(* IEC 61131-3 sources: codesys/project-view/Device/Plc Logic/Application/00-封装FC/DATA类型转换, 14 files *)

(* ---- FC_1DINT_TO_1DWORD.st ---- *)
FUNCTION FC_1DINT_TO_1DWORD : DWORD
VAR_INPUT
	diIN:DINT;
END_VAR
VAR
	pdw:POINTER TO DWORD;
END_VAR
// --- implementation ---
pdw:=ADR(diIN);
FC_1DINT_TO_1DWORD:=pdw^;
END_FUNCTION

(* ---- FC_1DWORD_TO_1REAL.st ---- *)
FUNCTION FC_1DWORD_TO_1REAL : REAL
VAR_INPUT
	dwIN:DWORD;
END_VAR
VAR
	pr:POINTER TO REAL;
END_VAR
// --- implementation ---
pr:=ADR(dwIN);
FC_1DWORD_TO_1REAL:=pr^;
END_FUNCTION

(* ---- FC_1REAL_TO_1DWORD.st ---- *)
FUNCTION FC_1REAL_TO_1DWORD : DWORD
VAR_INPUT
	rIN:DWORD;
END_VAR
VAR
	pdw:POINTER TO DWORD;
END_VAR
// --- implementation ---
pdw:=ADR(rIN);
FC_1REAL_TO_1DWORD:=pdw^;
END_FUNCTION

(* ---- FC_1REAL_TO_2WORD.st ---- *)
FUNCTION FC_1REAL_TO_2WORD : BOOL
VAR_INPUT
	rIN:REAL;
END_VAR
VAR_OUTPUT
	wOUT0:WORD;
	wOUT1:WORD;
END_VAR
VAR
	dw:DWORD;
	pdw:POINTER TO DWORD;
END_VAR
// --- implementation ---
pdw:=ADR(rIN);
dw:=pdw^;
wOUT0:=DWORD_TO_WORD(SHR(dw,0));
wOUT1:=DWORD_TO_WORD(SHR(dw,16));
FC_1REAL_TO_2WORD:=TRUE;
END_FUNCTION

(* ---- FC_1REAL_TO_4BYTE.st ---- *)
FUNCTION FC_1REAL_TO_4BYTE : BOOL
VAR_INPUT
	rIN:REAL;
END_VAR
VAR_OUTPUT
	byOUT0:BYTE;
	byOUT1:BYTE;
	byOUT2:BYTE;
	byOUT3:BYTE;
END_VAR
VAR
	dw:DWORD;
	pdw:POINTER TO DWORD;
END_VAR
// --- implementation ---
pdw:=ADR(rIN);
dw:=pdw^;
byOUT0:=DWORD_TO_BYTE(SHR(dw,0));
byOUT1:=DWORD_TO_BYTE(SHR(dw,8));
byOUT2:=DWORD_TO_BYTE(SHR(dw,16));
byOUT3:=DWORD_TO_BYTE(SHR(dw,24));
FC_1REAL_TO_4BYTE :=TRUE;
END_FUNCTION

(* ---- FC_1WORD_TO_2BYTE.st ---- *)
FUNCTION FC_1WORD_TO_2BYTE :BOOL
VAR_INPUT
	wIN:WORD;
END_VAR
VAR_OUTPUT
	byOUT0:BYTE;
	byOUT1:BYTE;
END_VAR
// --- implementation ---
byOUT0:=WORD_TO_BYTE(SHR(wIN,0));
byOUT1:=WORD_TO_BYTE(SHR(wIN,8));
END_FUNCTION

(* ---- FC_1WORD_TO_ARR16BOOL.st ---- *)
FUNCTION FC_1WORD_TO_ARR16BOOL : ARRAY [0..15] OF BOOL
VAR_INPUT
	wIN:WORD;
END_VAR
VAR
END_VAR
// --- implementation ---
FC_1WORD_TO_ARR16BOOL[0]:=TO_BOOL(wIN.0);
FC_1WORD_TO_ARR16BOOL[1]:=TO_BOOL(wIN.1);
FC_1WORD_TO_ARR16BOOL[2]:=TO_BOOL(wIN.2);
FC_1WORD_TO_ARR16BOOL[3]:=TO_BOOL(wIN.3);
FC_1WORD_TO_ARR16BOOL[4]:=TO_BOOL(wIN.4);
FC_1WORD_TO_ARR16BOOL[5]:=TO_BOOL(wIN.5);
FC_1WORD_TO_ARR16BOOL[6]:=TO_BOOL(wIN.6);
FC_1WORD_TO_ARR16BOOL[7]:=TO_BOOL(wIN.7);
FC_1WORD_TO_ARR16BOOL[8]:=TO_BOOL(wIN.8);
FC_1WORD_TO_ARR16BOOL[9]:=TO_BOOL(wIN.9);
FC_1WORD_TO_ARR16BOOL[10]:=TO_BOOL(wIN.10);
FC_1WORD_TO_ARR16BOOL[11]:=TO_BOOL(wIN.11);
FC_1WORD_TO_ARR16BOOL[12]:=TO_BOOL(wIN.12);
FC_1WORD_TO_ARR16BOOL[13]:=TO_BOOL(wIN.13);
FC_1WORD_TO_ARR16BOOL[14]:=TO_BOOL(wIN.14);
FC_1WORD_TO_ARR16BOOL[15]:=TO_BOOL(wIN.15);
END_FUNCTION

(* ---- FC_1WORD_TO_ARR16WORD.st ---- *)
FUNCTION FC_1WORD_TO_ARR16WORD : ARRAY [0..15] OF WORD
VAR_INPUT
	wIN:WORD;
END_VAR
VAR
END_VAR
// --- implementation ---
FC_1WORD_TO_ARR16WORD[0]:=TO_WORD(wIN.0);
FC_1WORD_TO_ARR16WORD[1]:=TO_WORD(wIN.1);
FC_1WORD_TO_ARR16WORD[2]:=TO_WORD(wIN.2);
FC_1WORD_TO_ARR16WORD[3]:=TO_WORD(wIN.3);
FC_1WORD_TO_ARR16WORD[4]:=TO_WORD(wIN.4);
FC_1WORD_TO_ARR16WORD[5]:=TO_WORD(wIN.5);
FC_1WORD_TO_ARR16WORD[6]:=TO_WORD(wIN.6);
FC_1WORD_TO_ARR16WORD[7]:=TO_WORD(wIN.7);
FC_1WORD_TO_ARR16WORD[8]:=TO_WORD(wIN.8);
FC_1WORD_TO_ARR16WORD[9]:=TO_WORD(wIN.9);
FC_1WORD_TO_ARR16WORD[10]:=TO_WORD(wIN.10);
FC_1WORD_TO_ARR16WORD[11]:=TO_WORD(wIN.11);
FC_1WORD_TO_ARR16WORD[12]:=TO_WORD(wIN.12);
FC_1WORD_TO_ARR16WORD[13]:=TO_WORD(wIN.13);
FC_1WORD_TO_ARR16WORD[14]:=TO_WORD(wIN.14);
FC_1WORD_TO_ARR16WORD[15]:=TO_WORD(wIN.15);
END_FUNCTION

(* ---- FC_2BYTE_TO_1WORD.st ---- *)
FUNCTION FC_2BYTE_TO_1WORD : WORD
VAR_INPUT
	byIN0:BYTE;
	byIN1:BYTE;
END_VAR
VAR
	w:WORD;
END_VAR
// --- implementation ---
w:=SHL(BYTE_TO_WORD(byIN1),8)+SHL(BYTE_TO_WORD(byIN0),0);
FC_2BYTE_TO_1WORD:=w;
END_FUNCTION

(* ---- FC_2UINT_TO_1REAL.st ---- *)
FUNCTION FC_2UINT_TO_1REAL : REAL
VAR_INPUT
	uiIN0:UINT;
	uiIN1:UINT;
END_VAR
VAR
	dui:UDINT;
	pr:POINTER TO REAL;
END_VAR
// --- implementation ---
dui:=SHL(WORD_TO_DWORD(uiIN1),16)+SHL(WORD_TO_DWORD(uiIN0),0);
pr:=ADR(dui);
FC_2UINT_TO_1REAL:=pr^;
END_FUNCTION

(* ---- FC_2WORD_TO_1REAL.st ---- *)
FUNCTION FC_2WORD_TO_1REAL : REAL
VAR_INPUT
	wIN0:WORD;
	wIN1:WORD;
END_VAR
VAR
	dw:DWORD;
	pr:POINTER TO REAL;
END_VAR
// --- implementation ---
dw:=SHL(WORD_TO_DWORD(wIN1),16)+SHL(WORD_TO_DWORD(wIN0),0);
pr:=ADR(dw);
FC_2WORD_TO_1REAL:=pr^;
END_FUNCTION

(* ---- FC_4BYTE_TO_1REAL.st ---- *)
FUNCTION FC_4BYTE_TO_1REAL : REAL
VAR_INPUT
	byIN0:BYTE;
	byIN1:BYTE;
	byIN2:BYTE;
	byIN3:BYTE;
END_VAR
VAR
	dw:DWORD;
	pr:POINTER TO REAL;
END_VAR
// --- implementation ---
dw:=SHL(BYTE_TO_DWORD(byIN3),24)+SHL(BYTE_TO_DWORD(byIN2),16)+SHL(BYTE_TO_DWORD(byIN1),8)+SHL(BYTE_TO_DWORD(byIN0),0);
pr:=ADR(dw);
FC_4BYTE_TO_1REAL:=pr^;
END_FUNCTION

(* ---- FC_ARR16BOOL_TO_1WORD.st ---- *)
FUNCTION FC_ARR16BOOL_TO_1WORD : WORD
VAR_INPUT
	axIN:ARRAY [0..15] OF BOOL;
END_VAR
VAR
END_VAR
// --- implementation ---
FC_ARR16BOOL_TO_1WORD.0:=TO_BIT(axIN[0]);
FC_ARR16BOOL_TO_1WORD.1:=TO_BIT(axIN[1]);
FC_ARR16BOOL_TO_1WORD.2:=TO_BIT(axIN[2]);
FC_ARR16BOOL_TO_1WORD.3:=TO_BIT(axIN[3]);
FC_ARR16BOOL_TO_1WORD.4:=TO_BIT(axIN[4]);
FC_ARR16BOOL_TO_1WORD.5:=TO_BIT(axIN[5]);
FC_ARR16BOOL_TO_1WORD.6:=TO_BIT(axIN[6]);
FC_ARR16BOOL_TO_1WORD.7:=TO_BIT(axIN[7]);
FC_ARR16BOOL_TO_1WORD.8:=TO_BIT(axIN[8]);
FC_ARR16BOOL_TO_1WORD.9:=TO_BIT(axIN[9]);
FC_ARR16BOOL_TO_1WORD.10:=TO_BIT(axIN[10]);
FC_ARR16BOOL_TO_1WORD.11:=TO_BIT(axIN[11]);
FC_ARR16BOOL_TO_1WORD.12:=TO_BIT(axIN[12]);
FC_ARR16BOOL_TO_1WORD.13:=TO_BIT(axIN[13]);
FC_ARR16BOOL_TO_1WORD.14:=TO_BIT(axIN[14]);
FC_ARR16BOOL_TO_1WORD.15:=TO_BIT(axIN[15]);
END_FUNCTION

(* ---- FC_ARR16WORD_TO_1WORD.st ---- *)
FUNCTION FC_ARR16WORD_TO_1WORD : WORD
VAR_INPUT
	awIN:ARRAY [0..15] OF WORD;
END_VAR
VAR
END_VAR
// --- implementation ---
FC_ARR16WORD_TO_1WORD[0]:=TO_WORD(awIN[0]);
FC_ARR16WORD_TO_1WORD[1]:=TO_WORD(awIN[1]);
FC_ARR16WORD_TO_1WORD[2]:=TO_WORD(awIN[2]);
FC_ARR16WORD_TO_1WORD[3]:=TO_WORD(awIN[3]);
FC_ARR16WORD_TO_1WORD[4]:=TO_WORD(awIN[4]);
FC_ARR16WORD_TO_1WORD[5]:=TO_WORD(awIN[5]);
FC_ARR16WORD_TO_1WORD[6]:=TO_WORD(awIN[6]);
FC_ARR16WORD_TO_1WORD[7]:=TO_WORD(awIN[7]);
FC_ARR16WORD_TO_1WORD[8]:=TO_WORD(awIN[8]);
FC_ARR16WORD_TO_1WORD[9]:=TO_WORD(awIN[9]);
FC_ARR16WORD_TO_1WORD[10]:=TO_WORD(awIN[10]);
FC_ARR16WORD_TO_1WORD[11]:=TO_WORD(awIN[11]);
FC_ARR16WORD_TO_1WORD[12]:=TO_WORD(awIN[12]);
FC_ARR16WORD_TO_1WORD[13]:=TO_WORD(awIN[13]);
FC_ARR16WORD_TO_1WORD[14]:=TO_WORD(awIN[14]);
FC_ARR16WORD_TO_1WORD[15]:=TO_WORD(awIN[15]);
END_FUNCTION
